// TIA Portal V20 export
// export: Created 2026-10-19T18:06:58.9116325Z, ExportSetting WithDefaults, DisplayName Totally Integrated Automation Portal, DisplayVersion V20 Update 6, DisplayName TIA Portal Openness, DisplayVersion V20 Update 6, DisplayName TIA Portal Version Control Interface, DisplayVersion V20 Update 6, DisplayName SINAMICS Startdrive Advanced, DisplayVersion V20 SP1, DisplayName SINAMICS Startdrive G130, G150, S120, S150, SINAMICS MV, G220, S200, S210, DisplayVersion V20 SP1, DisplayName SINAMICS Startdrive G110M, G120, G120C, G120D, G120P, G115D, DisplayVersion V20 SP1, DisplayName STEP 7 Professional, DisplayVersion V20 Update 6, DisplayName STEP 7 Safety, DisplayVersion V20 Update 2, DisplayName WinCC Basic/Comfort/Advanced, DisplayVersion V20 Update 6, DisplayName WinCC Unified, DisplayVersion V20 Update 6
DATA_BLOCK "MB_Device_Status"   // DB119
{ S7_Optimized_Access := 'TRUE' }
VERSION : 0.1
// stored: AutoNumber true, DBAccessibleFromOPCUA true, DBAccessibleFromWebserver true, InstanceOfName SAI_MB_DeviceStatus, InstanceOfType UDT, IsOnlyStoredInLoadMemory false, IsWriteProtectedInAS false
"SAI_MB_DeviceStatus"
   // VAR
   //    "Alternate weight unit" : Bool;
   //    "Run flat" : Bool;
   //    "Device specific bit 2" : Bool;
   //    "Device specific bit 3" : Bool;
   //    "Device specific bit 4" : Bool;
   //    "Device specific bit 5" : Bool;
   //    "Device specific bit 6" : Bool;
   //    "Device specific bit 7" : Bool;
   //    "Sequence bit 0" : Bool;
   //    "Sequence bit 1" : Bool;
   //    "Heart Beat" : Bool;
   //    "Data OK" : Bool;
   //    "Alarm Condition" : Bool;
   //    "Center of Zero" : Bool;
   //    Motion : Bool;
   //    "Net Mode" : Bool;
   // END_VAR
BEGIN
END_DATA_BLOCK
